Fanuc KAREL source: KT00757.KL

PROGRAM KT00757
%NOLOCKGROUP
VAR
  B1: BOOLEAN
  B2: BOOLEAN
  OUT: REAL
BEGIN
  B1 = TRUE
  B2 = FALSE
  B1 = TRUE
  B2 = FALSE
  OUT = ABS(B1)
END KT00757
